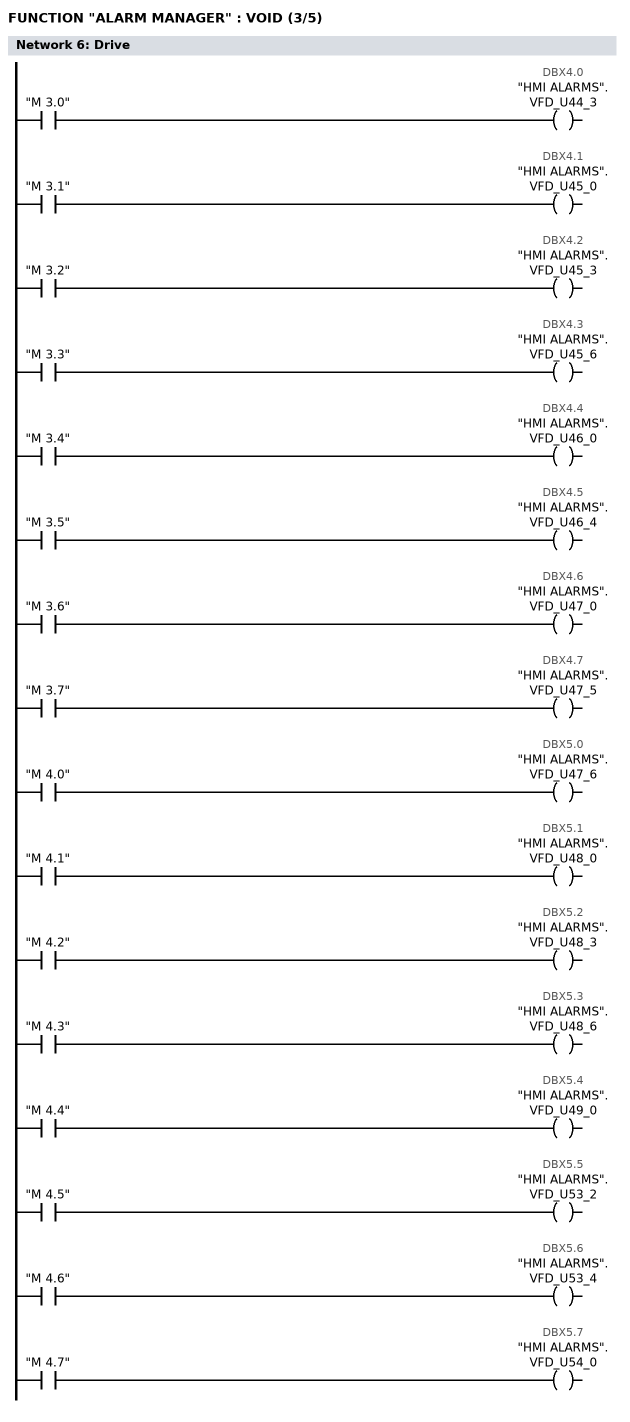

      A     "M 3.0";
      =     "HMI ALARMS".VFD_U44_3; // DBX4.0
//;
      A     "M 3.1";
      =     "HMI ALARMS".VFD_U45_0; // DBX4.1
//;
      A     "M 3.2";
      =     "HMI ALARMS".VFD_U45_3; // DBX4.2
//;
      A     "M 3.3";
      =     "HMI ALARMS".VFD_U45_6; // DBX4.3
//;
      A     "M 3.4";
      =     "HMI ALARMS".VFD_U46_0; // DBX4.4
//;
      A     "M 3.5";
      =     "HMI ALARMS".VFD_U46_4; // DBX4.5
//;
      A     "M 3.6";
      =     "HMI ALARMS".VFD_U47_0; // DBX4.6
//;
      A     "M 3.7";
      =     "HMI ALARMS".VFD_U47_5; // DBX4.7
//;
      A     "M 4.0";
      =     "HMI ALARMS".VFD_U47_6; // DBX5.0
//;
      A     "M 4.1";
      =     "HMI ALARMS".VFD_U48_0; // DBX5.1
//;
      A     "M 4.2";
      =     "HMI ALARMS".VFD_U48_3; // DBX5.2
//;
      A     "M 4.3";
      =     "HMI ALARMS".VFD_U48_6; // DBX5.3
//;
      A     "M 4.4";
      =     "HMI ALARMS".VFD_U49_0; // DBX5.4
//;
      A     "M 4.5";
      =     "HMI ALARMS".VFD_U53_2; // DBX5.5
//;
      A     "M 4.6";
      =     "HMI ALARMS".VFD_U53_4; // DBX5.6
//;
      A     "M 4.7";
      =     "HMI ALARMS".VFD_U54_0; // DBX5.7
NETWORK
TITLE =Sensor
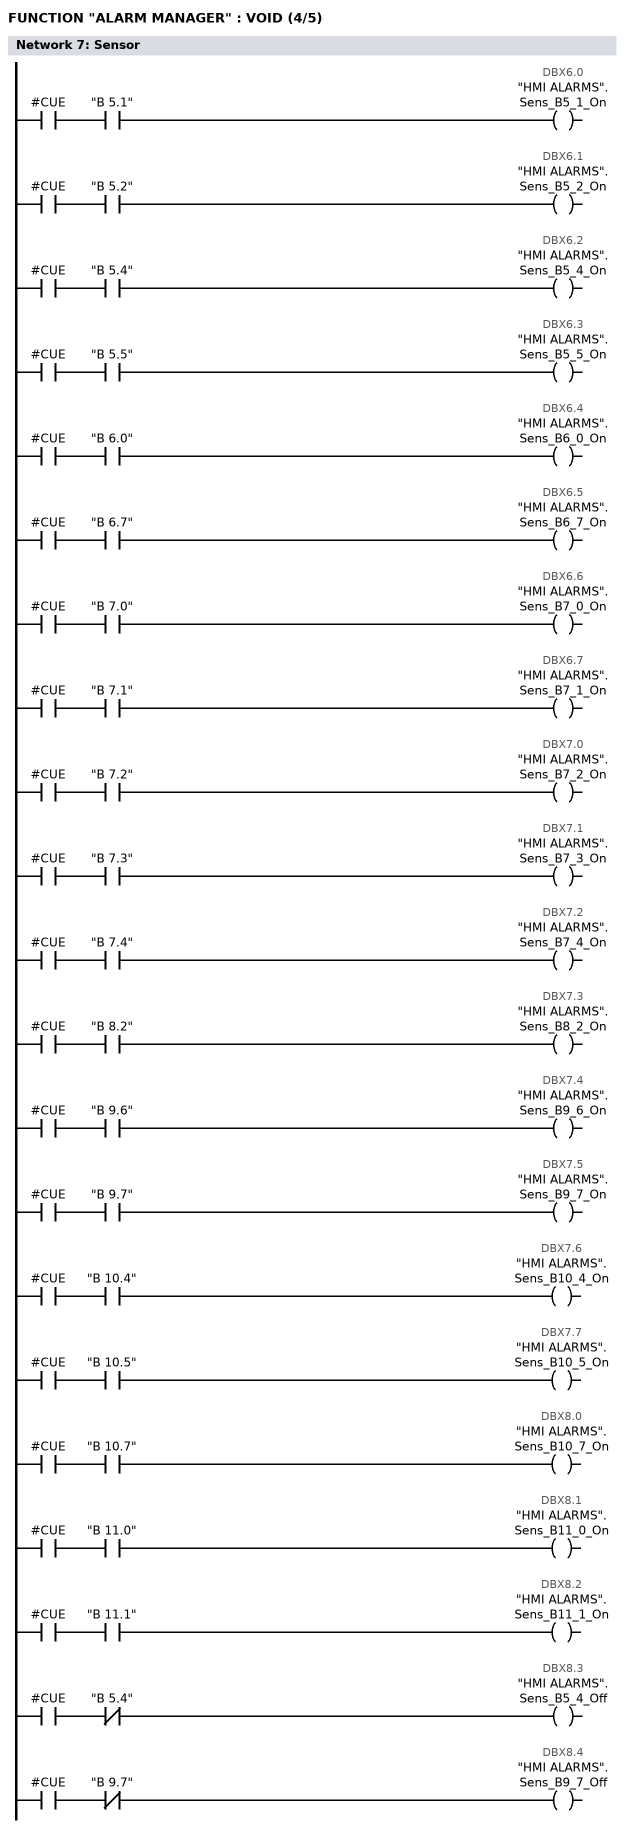

      A     #CUE;
      A     "B 5.1";
      =     "HMI ALARMS".Sens_B5_1_On; // DBX6.0
//;
      A     #CUE;
      A     "B 5.2";
      =     "HMI ALARMS".Sens_B5_2_On; // DBX6.1
//;
      A     #CUE;
      A     "B 5.4";
      =     "HMI ALARMS".Sens_B5_4_On; // DBX6.2
//;
      A     #CUE;
      A     "B 5.5";
      =     "HMI ALARMS".Sens_B5_5_On; // DBX6.3
//;
      A     #CUE;
      A     "B 6.0";
      =     "HMI ALARMS".Sens_B6_0_On; // DBX6.4
//;
      A     #CUE;
      A     "B 6.7";
      =     "HMI ALARMS".Sens_B6_7_On; // DBX6.5
//;
      A     #CUE;
      A     "B 7.0";
      =     "HMI ALARMS".Sens_B7_0_On; // DBX6.6
//;
      A     #CUE;
      A     "B 7.1";
      =     "HMI ALARMS".Sens_B7_1_On; // DBX6.7
//;
      A     #CUE;
      A     "B 7.2";
      =     "HMI ALARMS".Sens_B7_2_On; // DBX7.0
//;
      A     #CUE;
      A     "B 7.3";
      =     "HMI ALARMS".Sens_B7_3_On; // DBX7.1
//;
      A     #CUE;
      A     "B 7.4";
      =     "HMI ALARMS".Sens_B7_4_On; // DBX7.2
//;
      A     #CUE;
      A     "B 8.2";
      =     "HMI ALARMS".Sens_B8_2_On; // DBX7.3
//;
      A     #CUE;
      A     "B 9.6";
      =     "HMI ALARMS".Sens_B9_6_On; // DBX7.4
//;
      A     #CUE;
      A     "B 9.7";
      =     "HMI ALARMS".Sens_B9_7_On; // DBX7.5
//;
      A     #CUE;
      A     "B 10.4";
      =     "HMI ALARMS".Sens_B10_4_On; // DBX7.6
//;
      A     #CUE;
      A     "B 10.5";
      =     "HMI ALARMS".Sens_B10_5_On; // DBX7.7
//;
      A     #CUE;
      A     "B 10.7";
      =     "HMI ALARMS".Sens_B10_7_On; // DBX8.0
//;
      A     #CUE;
      A     "B 11.0";
      =     "HMI ALARMS".Sens_B11_0_On; // DBX8.1
//;
      A     #CUE;
      A     "B 11.1";
      =     "HMI ALARMS".Sens_B11_1_On; // DBX8.2
//;
      A     #CUE;
      AN    "B 5.4";
      =     "HMI ALARMS".Sens_B5_4_Off; // DBX8.3
//;
      A     #CUE;
      AN    "B 9.7";
      =     "HMI ALARMS".Sens_B9_7_Off; // DBX8.4
NETWORK
TITLE =Status
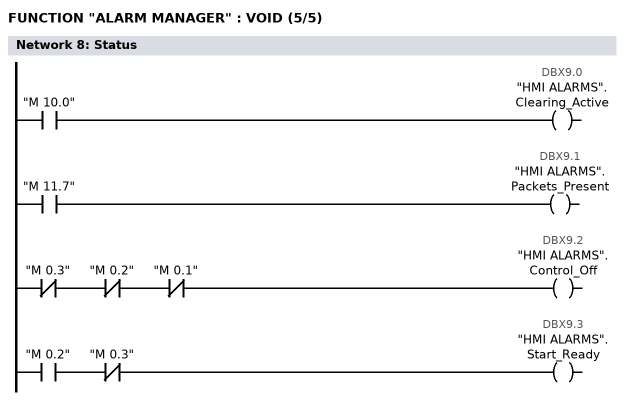

      A     "M 10.0";
      =     "HMI ALARMS".Clearing_Active; // DBX9.0
//;
      A     "M 11.7";
      =     "HMI ALARMS".Packets_Present; // DBX9.1
//;
      AN    "M 0.3";
      AN    "M 0.2";
      AN    "M 0.1";
      =     "HMI ALARMS".Control_Off; // DBX9.2
//;
      A     "M 0.2";
      AN    "M 0.3";
      =     "HMI ALARMS".Start_Ready; // DBX9.3
NETWORK
TITLE =Any Fault / Any Alarm - NS12 Alarm Bar (Control Flag)
//Bytes 0...8 = faults (spare bits are never set). Byte 9 bits 0...3 = status.
      A(    ;
      L     DB13.DBD    0; // Bytes 0...3
      L     L#0;
      <>D   ;
      )     ;
      O(    ;
      L     DB13.DBD    4; // Bytes 4...7
      L     L#0;
      <>D   ;
      )     ;
      O(    ;
      L     DB13.DBB    8; // Byte 8
      L     0;
      <>I   ;
      )     ;
      =     "HMI ALARMS".Any_Fault; // DBX9.6
//;
      A(    ;
      L     DB13.DBB    9; // Status 9.0...9.3
      L     B#16#F;
      AW    ;
      L     0;
      <>I   ;
      )     ;
      O     "HMI ALARMS".Any_Fault;
      =     "HMI ALARMS".Any_Alarm; // DBX9.7
END_FUNCTION

FUNCTION "FM350 COUNTERS" : VOID
TITLE =Counters
//FM350-2 : Counter Module Added to measure Collator Conveyors 4 & 10 Filling
//Surface Left, and to measure Packets Length & Width in order to Fit the Most
//Packets Number onto the Respective Conveyor... May 22
VERSION : 0.1


VAR_TEMP
  ENCODER_STOP : BOOL ;
  RETURN_RD : INT ;	//Print Pulse Read Function Return
  PRESS_LENGTH_3 : WORD ;	//Slat Conveyor 3 - Surface per Packet
  PACKET_LENGTH_4 : WORD ;	//Collator Conveyor 4 - Packet Length
  HALF_PACKET_LENGTH_4 : WORD ;	//Collator Conveyor 4 - Packet Length - Half
  PACKET_LENGTH_HALF_4 : WORD ;	//Collator Conveyor 4 - Packet Length + Half
  SURFACE_LENGTH_LEFT_4 : WORD ;	//Collator Conveyor 4 - Surface Length Left
  QTY_MAX_4 : REAL ;
  PACKET_WIDTH_10 : WORD ;	//Collator Conveyor 10 - Packet Width
  HALF_PACKET_WIDTH_10 : WORD ;	//Collator Conveyor 10 - Packet Width - Half
  PACKET_WIDTH_HALF_10 : WORD ;	//Collator Conveyor 10 - Packet Width + Half
  SURFACE_LENGTH_LEFT_10 : WORD ;
  QTY_MAX_10 : WORD ;
END_VAR
BEGIN
NETWORK
TITLE =Call DB

      OPN   "FM350 DB";
      CALL "CNT2_CTR" (//Control the FM 350-2
           DB_NO                    := W#16#2);

NETWORK
TITLE =FM350-2 Address Resets

      A     "M 167.7";
      JNB   M677;
      L     W#16#140;
      T     DBW   12;
//;
      L     DW#16#A00;
      T     DBD   14;
//;
      R     "M 167.7";

M677: NOP   0;
NETWORK
TITLE =Read Counters Jobs
//FM350-2 :  Job 100 = Read Counter 0,1,2,3
//           Job 101 = Read Counter 4,5,6,7
//           Then Transfer to DB2
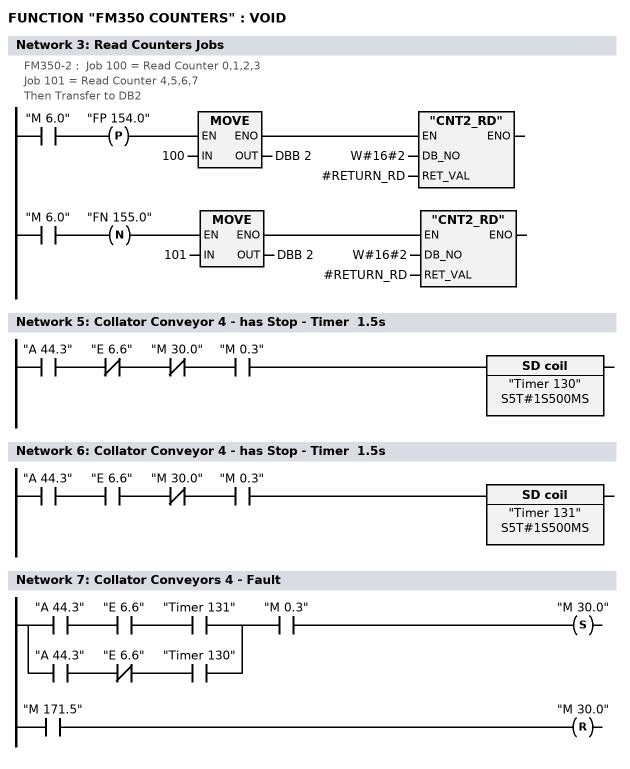
      A     "M 6.0";
      FP    "FP 154.0";
      JNB   M154;
      L     100;
      T     DBB    2;
      CALL "CNT2_RD" (
           DB_NO                    := W#16#2,
           RET_VAL                  := #RETURN_RD);

M154: NOP   0;

      A     "M 6.0";
      FN    "FN 155.0";
      JNB   M155;
      L     101;
      T     DBB    2;
      CALL "CNT2_RD" (
           DB_NO                    := W#16#2,
           RET_VAL                  := #RETURN_RD);

M155: NOP   0;
NETWORK
TITLE =
//Encoder Health Monitor


NETWORK
TITLE =Collator Conveyor 4 - has Stop - Timer  1.5s

      A     "A 44.3";
      AN    "E 6.6";
      AN    "M 30.0";
      A     "M 0.3";
      L     S5T#1S500MS;
      SD    "Timer 130";
NETWORK
TITLE =Collator Conveyor 4 - has Stop - Timer  1.5s

      A     "A 44.3";
      A     "E 6.6";
      AN    "M 30.0";
      A     "M 0.3";
      L     S5T#1S500MS;
      SD    "Timer 131";
NETWORK
TITLE =Collator Conveyors 4 - Fault

      A(    ;
      A     "A 44.3";
      A     "E 6.6";
      A     "Timer 131";
      O     ;
      A     "A 44.3";
      AN    "E 6.6";
      A     "Timer 130";
      )     ;
      A     "M 0.3";
      S     "M 30.0";
//;
      O     "M 171.5";
      R     "M 30.0";
NETWORK
TITLE =Collator Conveyors 4 - Lauer Comm

      OPN   "DB LAUER";

      A     "E 6.6";
      JC    M001;

      L     2#0;
      T     DBW  232;
      JU    M002;

M001: L     2#1;
      T     DBW  232;

M002: NOP   0;
END_FUNCTION

FUNCTION "ELEVATOR TEST FUNCTION" : VOID
TITLE =
VERSION : 0.1

BEGIN
NETWORK
TITLE =


      A     "A 63.0";
      JCN   M003;
      A     "A 63.3";
      JCN   M002;
      L     MW   950;
      L     1;
      -I    ;
      T     MW   950;
      JU    M001;
M002: L     MW   950;
      L     1;
      +I    ;
      T     MW   950;
M001: L     MW   950;
      L     200;
      <=I   ;
      =     M    930.1;
      L     MW   950;
      L     10;
      <=I   ;
      =     M    930.0;
      L     MW   950;
      L     800;
      >=I   ;
      =     M    930.2;
      L     MW   950;
      L     990;
      >=I   ;
      =     M    930.3;
M003: CLR   ;


END_FUNCTION

ORGANIZATION_BLOCK "CYCLIC"
TITLE =Main Cycle
//v0.1 2026-11-20: FC9xx switches read from DB111 (kept at power-off) instead of
//MB280...MB282. Bit layout unchanged: M280.0 = DB111.DBX0.0 ... M282.4 = DBX2.4.
//v0.2 2026-11-20: PIW test blocks: DB111.DBX2.5 FC925 (C3), 2.6 FC932 (C4), 2.7
//FC955 (C10).
//v0.3 2026-11-23: test switches removed. NEW blocks called directly (= v0.2 with
//all "TESTING DB" switches = 1): FC911...FC986 with FC925 / FC932 / FC955 (direct
//PIW) for C3 / C4 / C10. OLD FC1011...FC1086 and FC924 / FC931 / FC954 no longer
//called, "TESTING DB" (DB111) no longer read. Back: load OB1 v0.2.
//v1.0 2026-11-23: CALL FC1220 "HMI ALARMS FC" (NS12 alarm bits in DB13).
VERSION : 1.0


VAR_TEMP
  OB1_EV_CLASS : BYTE ;	//Bits 0-3 = 1 (Coming event), Bits 4-7 = 1 (Event class 1)
  OB1_SCAN_1 : BYTE ;	//1 (Cold restart scan 1 of OB 1), 3 (Scan 2-n of OB 1)
  OB1_PRIORITY : BYTE ;	//1 (Priority of 1 is lowest)
  OB1_OB_NUMBR : BYTE ;	//1 (Organization block 1, OB1)
  OB1_RESERVED_1 : BYTE ;	//Reserved for system
  OB1_RESERVED_2 : BYTE ;	//Reserved for system
  OB1_PREV_CYCLE : INT ;	//Cycle time of previous OB1 scan (milliseconds)
  OB1_MIN_CYCLE : INT ;	//Minimum cycle time of OB1 (milliseconds)
  OB1_MAX_CYCLE : INT ;	//Maximum cycle time of OB1 (milliseconds)
  OB1_DATE_TIME : DATE_AND_TIME ;	//Date and time OB1 started
END_VAR
BEGIN
NETWORK
TITLE =Scan Time
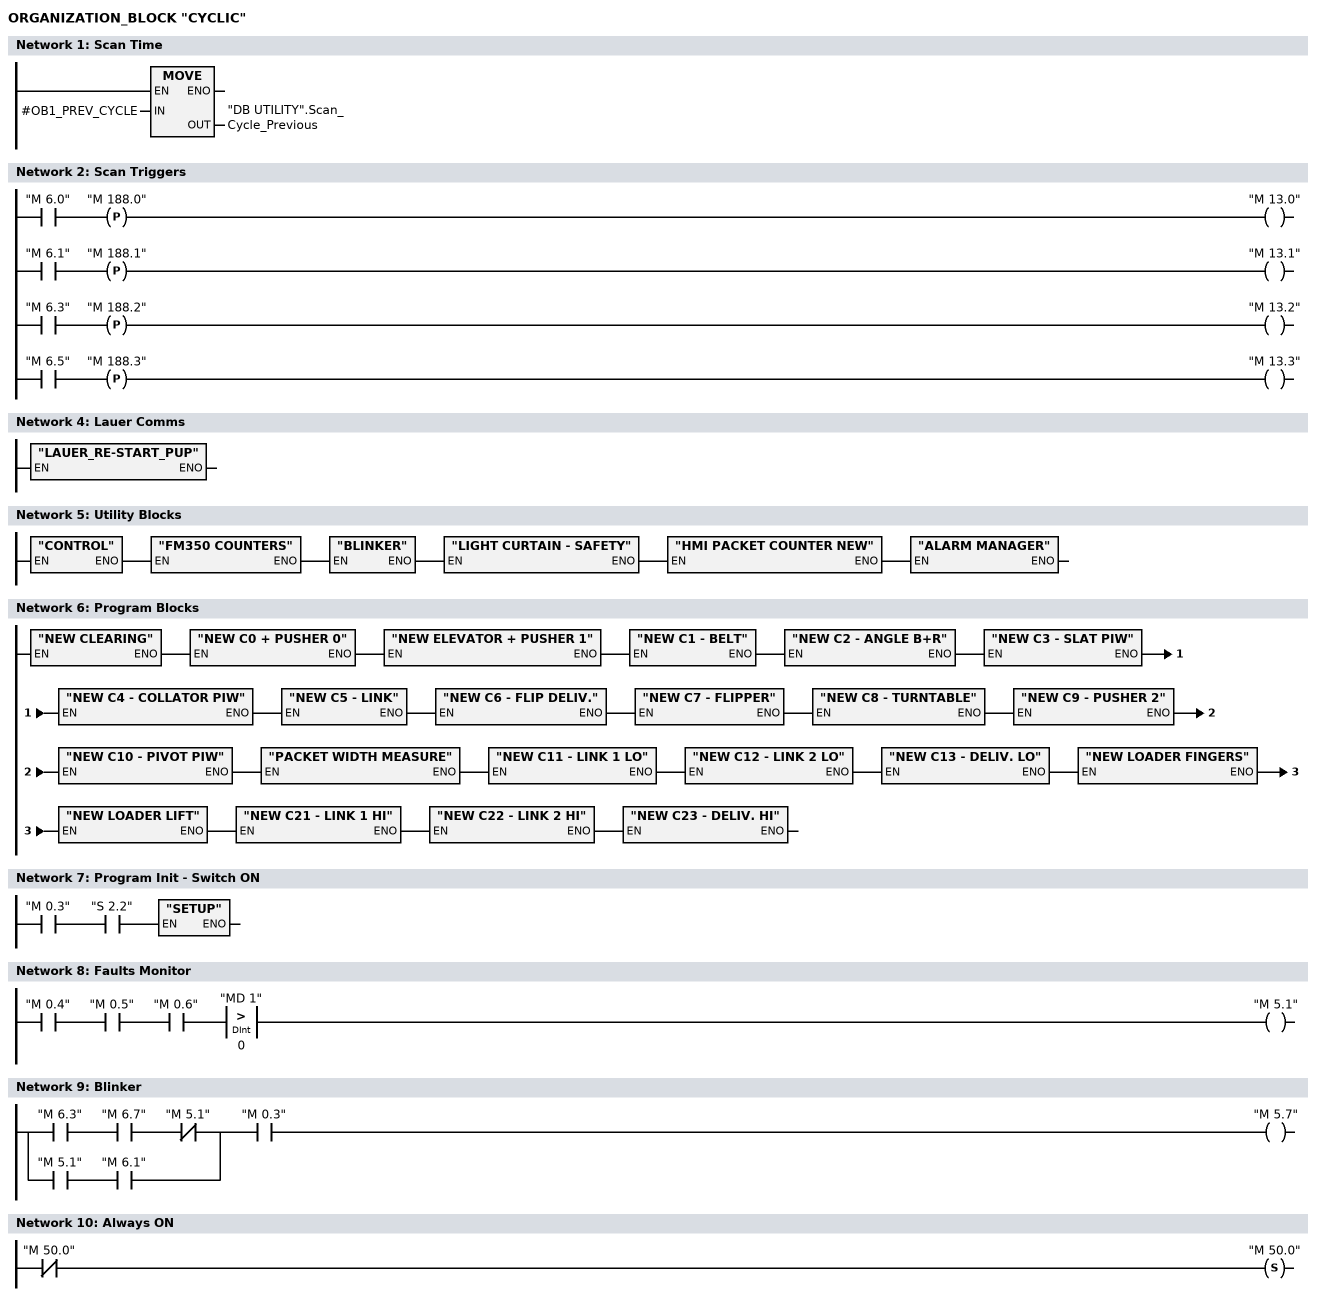

      L     #OB1_PREV_CYCLE;
      T     "DB UTILITY".Scan_Cycle_Previous;
NETWORK
TITLE =Scan Triggers

      A     "M 6.0";
      FP    "M 188.0";
      =     "M 13.0";
//;
      A     "M 6.1";
      FP    "M 188.1";
      =     "M 13.1";
//;
      A     "M 6.3";
      FP    "M 188.2";
      =     "M 13.2";
//;
      A     "M 6.5";
      FP    "M 188.3";
      =     "M 13.3";
NETWORK
TITLE =Packet Counters
//     CALL  "HMI PACKET COUNTER OLD"
//
//
//
//  CALL  "ELEVATOR TEST FUNCTION"
NETWORK
TITLE =Lauer Comms

      CALL "LAUER_RE-START_PUP" ;

NETWORK
TITLE =Utility Blocks

      CALL "CONTROL" ;
      CALL "FM350 COUNTERS" ;
      CALL "BLINKER" ;
      CALL "LIGHT CURTAIN - SAFETY" ;
      CALL "HMI PACKET COUNTER  NEW" ;
      CALL "ALARM MANAGER" ;// FC1220 - NS12 Alarm Bits (DB13)
NETWORK
TITLE =Program Blocks

      CALL "NEW CLEARING" ;// FC911
      CALL "NEW C0 + PUSHER 0" ;// FC912
      CALL "NEW ELEVATOR + PUSHER 1" ;// FC916
      CALL "NEW C1 - BELT" ;// FC918
      CALL "NEW C2 - ANGLE B+R" ;// FC922
      CALL "NEW C3 - SLAT PIW" ;// FC925 - PIW 328
      CALL "NEW C4 - COLLATOR PIW" ;// FC932 - PIW 330 / 332
      CALL "NEW C5 - LINK" ;// FC934
      CALL "NEW C6 - FLIP DELIV." ;// FC938
      CALL "NEW C7 - FLIPPER" ;// FC942
      CALL "NEW C8 - TURNTABLE" ;// FC948
      CALL "NEW C9 - PUSHER 2" ;// FC950
      CALL "NEW C10 - PIVOT PIW" ;// FC955 - PIW 334
      CALL "PACKET WIDTH MEASURE" ;// FC1210 - Width DB30 + Blanking DB31
      CALL "NEW C11 - LINK 1 LO" ;// FC958
      CALL "NEW C12 - LINK 2 LO" ;// FC962
      CALL "NEW C13 - DELIV. LO" ;// FC966
      CALL "NEW LOADER FINGERS" ;// FC970
      CALL "NEW LOADER LIFT" ;// FC974
      CALL "NEW C21 - LINK 1 HI" ;// FC978
      CALL "NEW C22 - LINK 2 HI" ;// FC982
      CALL "NEW C23 - DELIV. HI" ;// FC986


NETWORK
TITLE =Program Init - Switch ON

      A     "M 0.3";
      A     "S 2.2";
      JNB   M022;
      CALL "SETUP" ;

M022: NOP   0;
NETWORK
TITLE =Faults Monitor

      A     "M 0.4";
      A     "M 0.5";
      A     "M 0.6";
      A(    ;
      L     "MD 1";
      L     0;
      >D    ; // TODO later: <>D (MD1 < 0 when M 1.7 set) - kept as running
      )     ;
      =     "M 5.1";
NETWORK
TITLE =Blinker

      A(    ;
      A     "M 6.3";
      A     "M 6.7";
      AN    "M 5.1";
      O     ;
      A     "M 5.1";
      A     "M 6.1";
      )     ;
      A     "M 0.3";
      =     "M 5.7";
NETWORK
TITLE =Always ON

      AN    "M 50.0";
      S     "M 50.0";
END_ORGANIZATION_BLOCK

ORGANIZATION_BLOCK "Cyclic 100mS"
TITLE = "Cyclic Interrupt"
VERSION : 0.1


VAR_TEMP
  OB35_EV_CLASS : BYTE ;	//Bits 0-3 = 1 (Coming event), Bits 4-7 = 1 (Event class 1)
  OB35_STRT_INF : BYTE ;	//16#36 (OB 35 has started)
  OB35_PRIORITY : BYTE ;	//Priority of OB Execution
  OB35_OB_NUMBR : BYTE ;	//35 (Organization block 35, OB35)
  OB35_RESERVED_1 : BYTE ;	//Reserved for system
  OB35_RESERVED_2 : BYTE ;	//Reserved for system
  OB35_PHASE_OFFSET : WORD ;	//Phase offset (msec)
  OB35_RESERVED_3 : INT ;	//Reserved for system
  OB35_EXC_FREQ : INT ;	//Frequency of execution (msec)
  OB35_DATE_TIME : DATE_AND_TIME ;	//Date and time OB35 started
END_VAR
BEGIN
NETWORK
TITLE =CYCLIC 100 mS

      CALL "GENERAL FAULTS" ;
      CALL "HMI CONTROL" ;
      CALL "HMI COMMS" ;
      CALL "LIGHT BAR" ;

//  CALL  "Sensor Check Calls"
NETWORK
TITLE =Lauer Comms

      CALL "LAUER CALL" ;

NETWORK
TITLE =Lauer Comms

      CALL "LAUER COMM FC" (
           UBDB                     := "DB LAUER",
           RXFA                     := 36,
           RXLE                     := 32,
           TXFA                     := 3,
           TXLE                     := 32,
           RSET                     := "M 210.1",
           TIMT                     := T    105,
           TIMZ                     := S5T#1S,
           COFF                     := "LAUER RESTART FC",
           INIT                     := "LAUER COMM ERR FC",
           RFLM                     := "M 210.0",
           EROR                     := "M 210.2");
END_ORGANIZATION_BLOCK

ORGANIZATION_BLOCK "I/O_FLT1"
TITLE = "I/O Point Fault"
VERSION : 0.1


VAR_TEMP
  OB82_EV_CLASS : BYTE ;	//16#39, Event class 3, Entering event state, Internal fault event
  OB82_FLT_ID : BYTE ;	//16#XX, Fault identifcation code
  OB82_PRIORITY : BYTE ;	//Priority of OB Execution
  OB82_OB_NUMBR : BYTE ;	//82 (Organization block 82, OB82)
  OB82_RESERVED_1 : BYTE ;	//Reserved for system
  OB82_IO_FLAG : BYTE ;	//Input (01010100), Output (01010101)
  OB82_MDL_ADDR : WORD ;	//Base address of module with fault
  OB82_MDL_DEFECT : BOOL ;	//Module defective
  OB82_INT_FAULT : BOOL ;	//Internal fault
  OB82_EXT_FAULT : BOOL ;	//External fault
  OB82_PNT_INFO : BOOL ;	//Point information
  OB82_EXT_VOLTAGE : BOOL ;	//External voltage low
  OB82_FLD_CONNCTR : BOOL ;	//Field wiring connector missing
  OB82_NO_CONFIG : BOOL ;	//Module has no configuration data
  OB82_CONFIG_ERR : BOOL ;	//Module has configuration error
  OB82_MDL_TYPE : BYTE ;	//Type of module
  OB82_SUB_MDL_ERR : BOOL ;	//Sub-Module is missing or has error
  OB82_COMM_FAULT : BOOL ;	//Communication fault
  OB82_MDL_STOP : BOOL ;	//Module is stopped
  OB82_WTCH_DOG_FLT : BOOL ;	//Watch dog timer stopped module
  OB82_INT_PS_FLT : BOOL ;	//Internal power supply fault
  OB82_PRIM_BATT_FLT : BOOL ;	//Primary battery is in fault
  OB82_BCKUP_BATT_FLT : BOOL ;	//Backup battery is in fault
  OB82_RESERVED_2 : BOOL ;	//Reserved for system
  OB82_RACK_FLT : BOOL ;	//Rack fault, only for bus interface module
  OB82_PROC_FLT : BOOL ;	//Processor fault
  OB82_EPROM_FLT : BOOL ;	//EPROM fault
  OB82_RAM_FLT : BOOL ;	//RAM fault
  OB82_ADU_FLT : BOOL ;	//ADU fault
  OB82_FUSE_FLT : BOOL ;	//Fuse fault
  OB82_HW_INTR_FLT : BOOL ;	//Hardware interupt input in fault
  OB82_RESERVED_3 : BOOL ;	//Reserved for system
  OB82_DATE_TIME : DATE_AND_TIME ;	//Date and time OB82 started
END_VAR
BEGIN
NETWORK
TITLE =

END_ORGANIZATION_BLOCK

ORGANIZATION_BLOCK "RACK_FLT"
TITLE = "Loss Of Rack Fault"
VERSION : 0.1


VAR_TEMP
  OB86_EV_CLASS : BYTE ;	//16#38/39 Event class 3
  OB86_FLT_ID : BYTE ;	//16#C1/C4/C5, Fault identifcation code
  OB86_PRIORITY : BYTE ;	//Priority of OB Execution
  OB86_OB_NUMBR : BYTE ;	//86 (Organization block 86, OB86)
  OB86_RESERVED_1 : BYTE ;	//Reserved for system
  OB86_RESERVED_2 : BYTE ;	//Reserved for system
  OB86_MDL_ADDR : WORD ;	//Base address of IM module in rack with fault
  OB86_RACKS_FLTD : ARRAY  [0 .. 31 ] OF BOOL ;	//Racks in fault
  OB86_DATE_TIME : DATE_AND_TIME ;	//Date and time OB86 started
END_VAR
BEGIN
NETWORK
TITLE =

END_ORGANIZATION_BLOCK

ORGANIZATION_BLOCK "OB100"
TITLE =Start up    OB100
VERSION : 0.1


VAR_TEMP
  OB100_EV_CLASS : BYTE ;	//16#13, Event class 1, Entering event state, Event logged in diagnostic buffer
  OB100_STRTUP : BYTE ;	//16#81/82/83/84 Method of startup
  OB100_PRIORITY : BYTE ;	//27 (Priority of 1 is lowest)
  OB100_OB_NUMBR : BYTE ;	//100 (Organization block 100, OB100)
  OB100_RESERVED_1 : BYTE ;	//Reserved for system
  OB100_RESERVED_2 : BYTE ;	//Reserved for system
  OB100_STOP : WORD ;	//Event that caused CPU to stop (16#4xxx)
  OB100_STRT_INFO : DWORD ;	//Information on how system started
  OB100_DATE_TIME : DATE_AND_TIME ;	//Date and time OB100 started
END_VAR
BEGIN
NETWORK
TITLE =Lauer restart bit

      L     2#0; // Reset First cycle Flag
      =     "M 210.0";
NETWORK
TITLE =HMI On Lamp

      AN    "HMI_DB".TRANS_SYSTEM_RUN_STATUS;
      =     "HMI_DB".TRANS_SYSTEM_RUN_STATUS;
NETWORK
TITLE =DB Init

      R     "DEBOUNCER COUNTER DB".Conveyor_C3_Slat.FirstScan_Done;
      R     "DEBOUNCER COUNTER DB".Conveyor_C4_Collator.FirstScan_Done;
      R     "DEBOUNCER COUNTER DB".Conveyor_C5_Link.FirstScan_Done;
      R     "DEBOUNCER COUNTER DB".Conveyor_C6_Delivery.FirstScan_Done;
      R     "DEBOUNCER COUNTER DB".Conveyor_C10_Collator.FirstScan_Done;
      R     "DEBOUNCER COUNTER DB".Conveyor_C11_Link.FirstScan_Done;
      R     "DEBOUNCER COUNTER DB".Conveyor_C12_Link.FirstScan_Done;
      R     "DEBOUNCER COUNTER DB".Conveyor_C13_Delivery.FirstScan_Done;
      R     "DEBOUNCER COUNTER DB".Conveyor_C21_Link.FirstScan_Done;
      R     "DEBOUNCER COUNTER DB".Conveyor_C22_Link.FirstScan_Done;
      R     "DEBOUNCER COUNTER DB".Conveyor_C23_Delivery.FirstScan_Done;
END_ORGANIZATION_BLOCK

ORGANIZATION_BLOCK "PROG_ERR"
TITLE = "Programming Error"
VERSION : 0.1


VAR_TEMP
  OB121_EV_CLASS : BYTE ;	//16#25, Event class 2, Entering event state, Internal fault event
  OB121_SW_FLT : BYTE ;	//16#XX Software programming fault
  OB121_PRIORITY : BYTE ;	//Priority of OB Execution
  OB121_OB_NUMBR : BYTE ;	//121 (Organization block 121, OB121)
  OB121_BLK_TYPE : BYTE ;	//16#88/8A/8B/8C/8E Type of block fault occured in
  OB121_RESERVED_1 : BYTE ;	//Reserved for system
  OB121_FLT_REG : WORD ;	//16#XX Specific register that caused fault
  OB121_BLK_NUM : WORD ;	//Number of block that programming fault occured in
  OB121_PRG_ADDR : WORD ;	//Address in block where programming fault occured
  OB121_DATE_TIME : DATE_AND_TIME ;	//Date and time OB121 started
END_VAR
BEGIN
NETWORK
TITLE =

END_ORGANIZATION_BLOCK

ORGANIZATION_BLOCK "IO ACCESS_ERR"
TITLE = "Programming Error"
VERSION : 0.1


VAR_TEMP
  OB121_EV_CLASS : BYTE ;	//16#25, Event class 2, Entering event state, Internal fault event
  OB121_SW_FLT : BYTE ;	//16#XX Software programming fault
  OB121_PRIORITY : BYTE ;	//Priority of OB Execution
  OB121_OB_NUMBR : BYTE ;	//121 (Organization block 121, OB121)
  OB121_BLK_TYPE : BYTE ;	//16#88/8A/8B/8C/8E Type of block fault occured in
  OB121_RESERVED_1 : BYTE ;	//Reserved for system
  OB121_FLT_REG : WORD ;	//16#XX Specific register that caused fault
  OB121_BLK_NUM : WORD ;	//Number of block that programming fault occured in
  OB121_PRG_ADDR : WORD ;	//Address in block where programming fault occured
  OB121_DATE_TIME : DATE_AND_TIME ;	//Date and time OB121 started
END_VAR
BEGIN
NETWORK
TITLE =

END_ORGANIZATION_BLOCK

